FUNCTION_BLOCK StopPoint (* CAT Function Block Type *)
  (* Standard: 61499-2 *)
  (* Version 0.0, 11/22/2026, Schneider Electric, Lightweight stop point CAT *)
  PACKAGE Main;
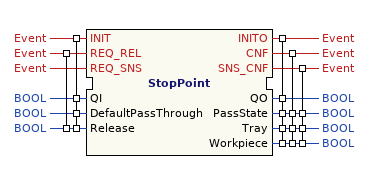
  EVENT_INPUT
    INIT WITH QI, DefaultPassThrough, Release; (* Initialization Request *)
    REQ_REL WITH Release; (* External release command update *)
    REQ_SNS; (* Request current tray and workpiece sensor states *)
  END_EVENT
  EVENT_OUTPUT
    INITO WITH QO, PassState, Tray, Workpiece; (* Initialization Confirm *)
    CNF WITH PassState, Tray, Workpiece; (* Pass-through state confirmation *)
    SNS_CNF WITH Tray, Workpiece, PassState; (* Tray or workpiece sensor update *)
  END_EVENT
  VAR_INPUT
    QI : BOOL := TRUE; (* Input event qualifier *)
    DefaultPassThrough : BOOL := FALSE; (* Startup mode (FALSE=Blocking/Up, TRUE=Pass-Through/Down) *)
    Release : BOOL := FALSE; (* External temporary release input *)
  END_VAR
  VAR_OUTPUT
    QO : BOOL; (* Output event qualifier *)
    PassState : BOOL; (* Effective pass-through state (TRUE=Down, FALSE=Up) *)
    Tray : BOOL; (* Tray present sensor state *)
    Workpiece : BOOL; (* Workpiece present sensor state *)
  END_VAR
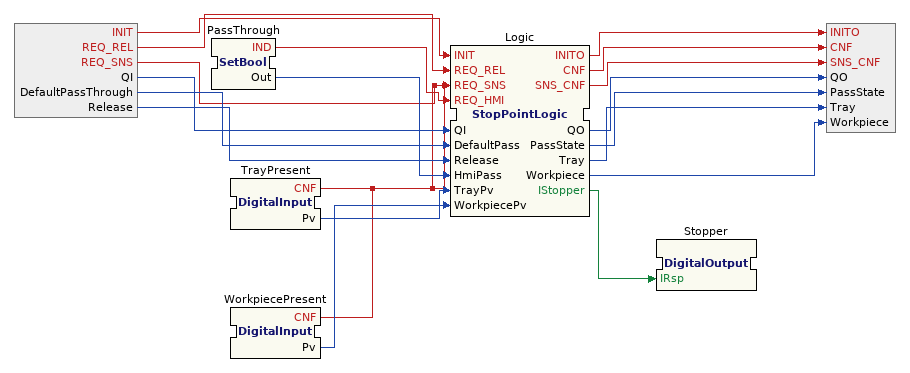
  FBS
    Stopper : DigitalOutput;
    TrayPresent : DigitalInput;
    WorkpiecePresent : DigitalInput;
    PassThrough : SetBool;
    Logic : StopPointLogic;
  END_FBS
  EVENT_CONNECTIONS
    INIT TO Logic.INIT;
    REQ_REL TO Logic.REQ_REL;
    REQ_SNS TO Logic.REQ_SNS;
    PassThrough.IND TO Logic.REQ_HMI;
    TrayPresent.CNF TO Logic.REQ_SNS;
    WorkpiecePresent.CNF TO Logic.REQ_SNS;
    Logic.INITO TO INITO;
    Logic.CNF TO CNF;
    Logic.SNS_CNF TO SNS_CNF;
  END_CONNECTIONS
  DATA_CONNECTIONS
    QI TO Logic.QI;
    DefaultPassThrough TO Logic.DefaultPass;
    Release TO Logic.Release;
    PassThrough.Out TO Logic.HmiPass;
    TrayPresent.Pv TO Logic.TrayPv;
    WorkpiecePresent.Pv TO Logic.WorkpiecePv;
    Logic.QO TO QO;
    Logic.PassState TO PassState;
    Logic.Tray TO Tray;
    Logic.Workpiece TO Workpiece;
  END_CONNECTIONS
  ADAPTER_CONNECTIONS
    Logic.IStopper TO Stopper.IRsp;
  END_CONNECTIONS
END_FUNCTION_BLOCK
